Fanuc KAREL source: kf00099.KL

-- PROVISIONAL review KL for V1013-1; original PC SHA256 bac3a317eaca79e310074db1165d5526428f9193d173e2386c2c05c1d7d807bb
-- Incomplete behavior may be omitted. Consult companion uncertainty JSON. Do not deploy.
PROGRAM KF00099
%NOLOCKGROUP
BEGIN
  -- UNRESOLVED_PC offsets 5-16; opcodes 2E,23
  -- UNRESOLVED_PC offsets 21-32; opcodes 2E,23
  -- UNRESOLVED_PC offsets 37-63; opcodes 27,27,9D,22,27,9D,31,7E,4A
  -- UNRESOLVED_PC offsets 68-72; opcodes 7F
END KF00099
